NAMESPACE TiaMcp_UnitA
DATA_BLOCK "TgpUnit_OperandDB"
{ S7_Optimized_Access := 'TRUE' }
VERSION : 0.1
NON_RETAIN
VAR
 Flag : Bool;
 Target : Bool;
END_VAR
BEGIN
END_DATA_BLOCK

END_NAMESPACE
